// TIA Portal V21 export
// export: Created 2026-11-08T19:47:41.2172749Z, ExportSetting WithDefaults, DisplayName Totally Integrated Automation Portal, DisplayVersion V21 Update 3, DisplayName STEP 7 Professional, DisplayVersion V21 Update 3, DisplayName STEP 7 Safety, DisplayVersion V21, DisplayName Tech WebApplication, DisplayVersion V21, DisplayName WinCC Basic/Comfort/Advanced, DisplayVersion V21 Update 3, DisplayName WinCC Unified, DisplayVersion V21 Update 3
FUNCTION "FC_Lad" : Void   // FC2, LAD
{ S7_Optimized_Access := 'TRUE' }
VERSION : 0.1
// stored: AutoNumber true, IsIECCheckEnabled false, SetENOAutomatically false, UDAEnableTagReadback false
   VAR_INPUT
      start : Bool;   // Start command
      "a" : Int;   // First addend
      "b" : Int;   // Second addend
   END_VAR
   VAR_OUTPUT
      running : Bool;   // Running state
      sum : Int;   // Sum of a and b
   END_VAR
BEGIN

REGION Network 1: Start latch
   // Copies the start command to the running state
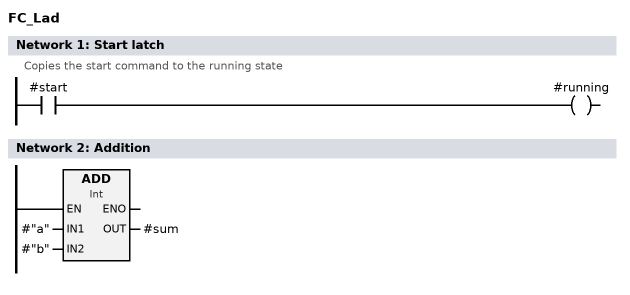
   RUNG wire#powerrail
      Contact( #start )
      Coil( #running )
   END_RUNG
   // the same network as SCL:
   #running := #start;
END_REGION

REGION Network 2: Addition
   RUNG wire#powerrail
      { S7_Templates := "SrcType := Int" } Add(in1 := #"a", in2 := #"b", out => #sum)
   END_RUNG
   // the same network as SCL:
   #sum := #"a" + #"b";
END_REGION
END_FUNCTION
